(* IEC 61131-3 sources: kns-port-domestic/targets/astra/src/POUs/Log/PRG_Slow, 2 files *)

(* ---- PRG_Slow.decl.st ---- *)
// Назначение: медленная задача (SlowTask): выгрузка снимка журнала в CSV по запросу MainTask
//             (GVL_Log.xExportReq). Запрос принимается, когда выгрузка не идёт, и снимается сразу после
//             публикации состояния Writing: MainTask ставит запрос только вне Writing, поэтому запись TRUE
//             из MainTask не теряется при вытеснении SlowTask (повторная команда до старта сливается с
//             первой). Число строк и код ошибки публикуются раньше состояния Done/Error: MainTask по
//             переходу состояния пишет событие с ними. Файловые операции не влияют на цикл логики (D-09).
// Автор:      kr0nsch
// Версия:     0.2.0
// Документ:   docs/DESIGN.md, разделы 4.3, 9.2
PROGRAM PRG_Slow
VAR
    fbCsv  : FB_EventLogCsv;        // выгрузка журнала
    xStart : BOOL;                  // запрос MainTask принят в этом цикле
END_VAR

(* ---- PRG_Slow.impl.st ---- *)
// запрос принимается, только пока выгрузка не идёт (фронт xExecute FB_EventLogCsv — по принятию)
xStart := GVL_Log.xExportReq AND fbCsv.eState <> E_LogExportState.Writing;
fbCsv(xExecute := xStart, sFileName := GVL_Const.LOG_CSV_FILE, fbLog := GVL_Log.fbEventLog);
// итог — до состояния: MainTask по переходу в Done/Error пишет событие с числом строк или кодом ошибки
IF fbCsv.xDone OR fbCsv.xError THEN
    GVL_Log.uiExportLines := fbCsv.uiLines;
    GVL_Log.udiExportError := fbCsv.udiError;
END_IF
GVL_Log.eExportState := fbCsv.eState;
// запрос снимается после публикации Writing: при Writing MainTask новый запрос не ставит
IF xStart THEN
    GVL_Log.xExportReq := FALSE;
END_IF
